// TIA Portal V21 export
// export: Created 2026-11-11T00:47:55.243187Z, ExportSetting WithDefaults, DisplayName Totally Integrated Automation Portal, DisplayVersion V21 Update 3, DisplayName STEP 7 Professional, DisplayVersion V21 Update 3, DisplayName STEP 7 Safety, DisplayVersion V21, DisplayName Tech WebApplication, DisplayVersion V21, DisplayName WinCC Basic/Comfort/Advanced, DisplayVersion V21 Update 3, DisplayName WinCC Unified, DisplayVersion V21 Update 3
FUNCTION_BLOCK "FB_Lad_ou021"   // FB347, LAD
{ S7_Optimized_Access := 'TRUE' }
VERSION : 0.1
// stored: AutoNumber true, IsIECCheckEnabled false, IsRetainMemResEnabled false, MemoryReserve 100, SetENOAutomatically false, UDAEnableTagReadback false
   VAR_INPUT
      v_req : Bool;
      v_interface : HW_INTERFACE;
      v_conf_data : Array[0..99] of Byte;
   END_VAR
   VAR_OUTPUT
      v_done : Bool;
      v_busy : Bool;
      v_error : Bool;
      v_status : DWord;
      v_err_loc : DWord;
   END_VAR
   VAR
      inst { S7_SetPoint := 'True'} : T_CONFIG;
   END_VAR
BEGIN

REGION Network 1: Description T_CONFIG
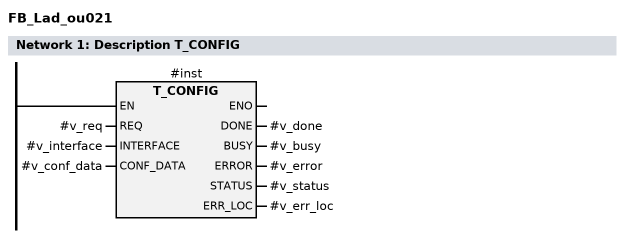
   RUNG wire#powerrail
      #inst.T_CONFIG(Req := #v_req, Interface := #v_interface, Conf_Data := #v_conf_data, Done => #v_done, Busy => #v_busy, Error => #v_error, Status => #v_status, Err_Loc => #v_err_loc)
   END_RUNG
   // the same network as SCL:
   #inst(Req := #v_req,   // T_CONFIG
         Interface := #v_interface,
         Conf_Data := #v_conf_data,
         Done => #v_done,
         Busy => #v_busy,
         Error => #v_error,
         Status => #v_status,
         Err_Loc => #v_err_loc);
END_REGION
END_FUNCTION_BLOCK
